{attribute 'qualified_only'}
VAR_GLOBAL
    // Display-only, not consumed by machine or safety permissives.
    stStatus : ST_EL6910Diagnostics;
END_VAR

(* stored: Version 1.1.0.1, ProductVersion 3.1.4026.18
   GVL GVL_EL6910Diagnostics: Id {78ef46cb-1437-4d1d-a484-74284eae251d} *)
